(* Logix 5000 project; controller R400_500_XLS vendor 1 type 14 code 216 rev 31.11; software revision 31.01; part 19 of 32 *)
(* tags used below, declared in another part *)
   Alarm : SINT;   // Wait 3 seconds
   Condenser : INT;
   DRYING : DINT;   // Drying id number
   FINAL_RINSE_MAX_NBR : INT;   // Maximum nimber of final rinse
   LowPressAlmSp : REAL;   // Pump pressure too low setpoint
   M : DINT[5];   // Memory Bits
   MaxTrtTempSp : REAL;
   ONS_FC85 : SINT;
   PURE_WATER_HEATING_TIME : DINT;   // Time before an alarm is thrown when the pure water tank is heating
   PWTnkTempAlmSp : REAL;   // Pure water tank temperature too high setpoint
   s00_Nb : STRING;
   s0_Nb : STRING;
   s2lastdigits : STRING;
   s36 : STRING;
   s360 : STRING;
   s3600 : STRING;
   s36000 : STRING;
   s360000 : STRING;
   s3600000 : STRING;
   s36000000 : STRING;
   s360000000 : STRING;
   sDigits1_2 : STRING;
   Service : DINT[2];   // Unused Service Mode Memory Bit
   ServicePassword : DINT;   // Service Password
   sInvertedPairs : STRING;
   sLastdigit : STRING;
   SRE3_Serial_Number : STRING;   // Serial number
   start_1 : SINT;
   start_2 : SINT;
   sTempo1 : STRING;
   sTempo2 : STRING;
   SumpTempAlmSp : REAL;   // Sump temperature too high setpoint
   Tmr : TIMER[107];
   bInibitAutologout : BOOL;   // Cancel AutoLogout
   BoilingValue : REAL;
   Cfg_10_Modules : BOOL;   // Chassis is configured 10 slots
   ChemicalName : STRING[9];   // Used by HMI
   COOLING_PHASE_TIME : DINT;   // Time of the cooling phase when time based drying
   DrainExtensionTime : DINT;
   iDelayBeforeFillingAuthAlarmMM : DINT;
   iDelayBeforeFillingAuthAlarmSS : DINT;
   iInactivityLogoutTime : DINT;   // Inactivity Logout Time In Minutes
   iInactivityPeriod : DINT;   // Inactivity Period before Logout * Value Must be greater than 0
   iPWClosingDelayMM : DINT;
   iPWClosingDelaySS : DINT;
   Non_Vented_with_Dry_Option : BOOL;
   NonVented_Without_Dry_Option : BOOL;
   NumInput : UDT_NUMERIC_INPUT[65];   // Numeric input
   NumInputReal : UDT_NUMERIC_INPUT_REAL[17];
   Screen_Ctrl : DINT;   // PLC Screen Request
   tDelayBeforeFillingAuthAlarm : TIMER;
   tDelayBeforeTankFillingAuthAlarm : TIMER;
   Tpb : DINT[11];
   tPureWaterTankClosingDelay : TIMER;
   tPWClosingDelay : TIMER;
   TRUE : BOOL;   // Always true bit
   Unit : Hrdwre;   // Unit Configuration
   Vented_with_Dry_Option : BOOL;
(* MainProgram, continued *)

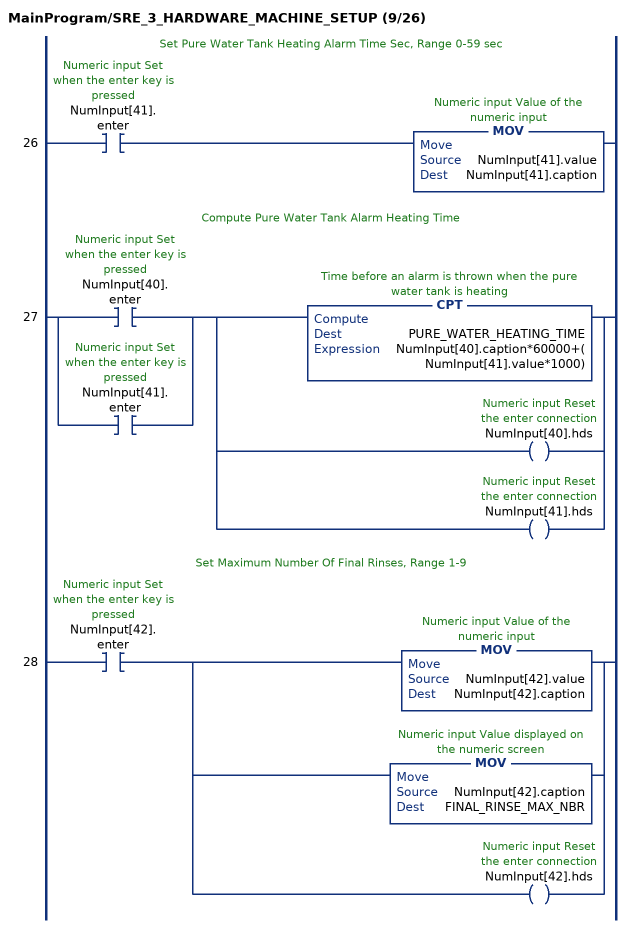
   [picture p363: MainProgram/SRE_3_HARDWARE_MACHINE_SETUP rungs 26-28]
   // Set Pure Water Tank Heating Alarm Time Sec, Range 0-59 sec
   26: XIC(NumInput[41].enter)MOV(NumInput[41].value,NumInput[41].caption);
   // Compute Pure Water Tank Alarm Heating Time
   27: [XIC(NumInput[40].enter) ,XIC(NumInput[41].enter) ][CPT(PURE_WATER_HEATING_TIME,NumInput[40].caption*60000+(NumInput[41].value*1000)) ,OTE(NumInput[40].hds) ,OTE(NumInput[41].hds) ];
   // Set Maximum Number Of Final Rinses, Range 1-9
   28: XIC(NumInput[42].enter)[MOV(NumInput[42].value,NumInput[42].caption) ,MOV(NumInput[42].caption,FINAL_RINSE_MAX_NBR) ,OTE(NumInput[42].hds) ];
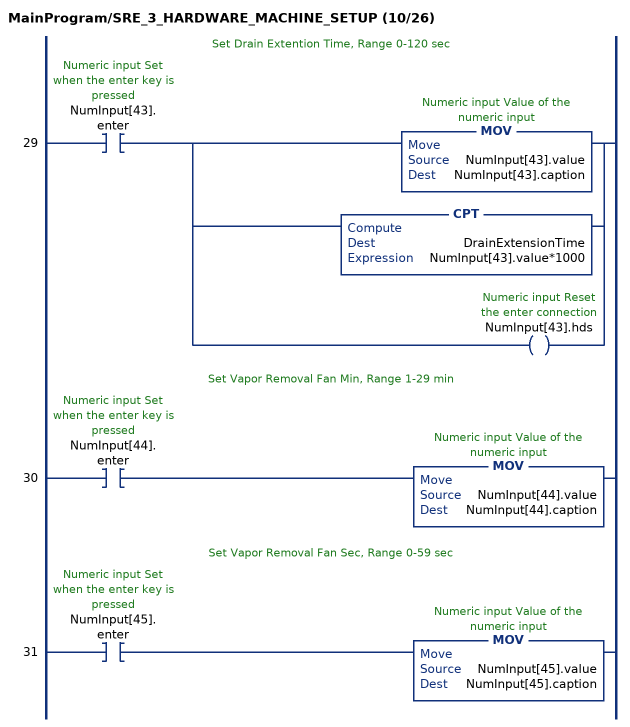
   // Set Drain Extention Time, Range 0-120 sec
   29: XIC(NumInput[43].enter)[MOV(NumInput[43].value,NumInput[43].caption) ,CPT(DrainExtensionTime,NumInput[43].value*1000) ,OTE(NumInput[43].hds) ];
   // Set Vapor Removal Fan Min, Range 1-29 min
   30: XIC(NumInput[44].enter)MOV(NumInput[44].value,NumInput[44].caption);
   // Set Vapor Removal Fan Sec, Range 0-59 sec
   31: XIC(NumInput[45].enter)MOV(NumInput[45].value,NumInput[45].caption);
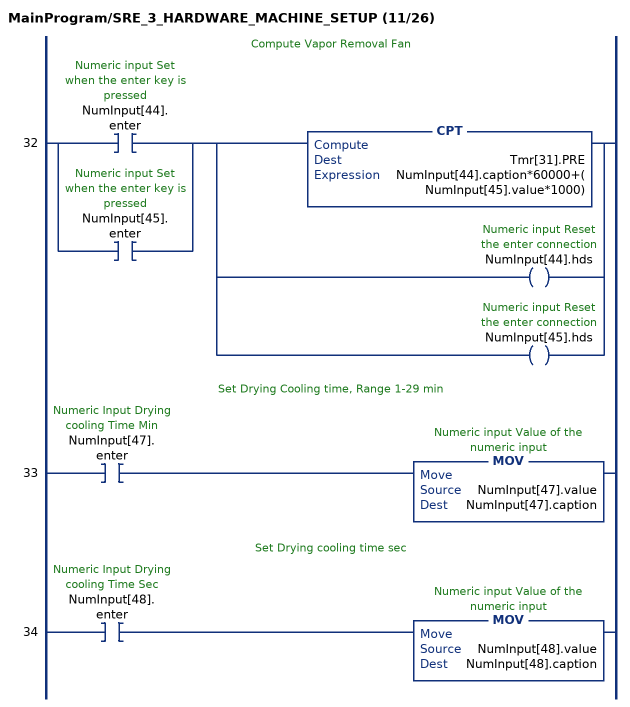
   // Compute Vapor Removal Fan
   32: [XIC(NumInput[44].enter) ,XIC(NumInput[45].enter) ][CPT(Tmr[31].PRE,NumInput[44].caption*60000+(NumInput[45].value*1000)) ,OTE(NumInput[44].hds) ,OTE(NumInput[45].hds) ];
   // Set Drying Cooling time, Range 1-29 min
   33: XIC(NumInput[47].enter)MOV(NumInput[47].value,NumInput[47].caption);
   // Set Drying cooling time sec
   34: XIC(NumInput[48].enter)MOV(NumInput[48].value,NumInput[48].caption);
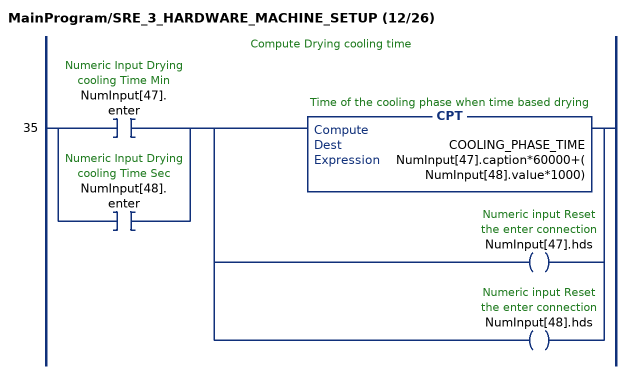
   // Compute Drying cooling time
   35: [XIC(NumInput[47].enter) ,XIC(NumInput[48].enter) ][CPT(COOLING_PHASE_TIME,NumInput[47].caption*60000+(NumInput[48].value*1000)) ,OTE(NumInput[47].hds) ,OTE(NumInput[48].hds) ];
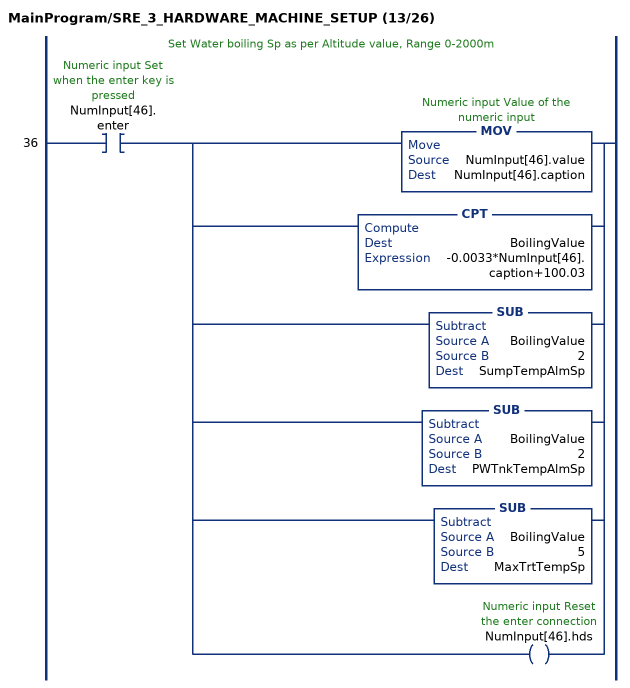
   // Set Water boiling Sp as per Altitude value, Range 0-2000m
   36: XIC(NumInput[46].enter)[MOV(NumInput[46].value,NumInput[46].caption) ,CPT(BoilingValue,-0.0033*NumInput[46].caption+100.03) ,SUB(BoilingValue,2,SumpTempAlmSp) ,SUB(BoilingValue,2,PWTnkTempAlmSp) ,SUB(BoilingValue,5,MaxTrtTempSp) ,OTE(NumInput[46].hds) ];
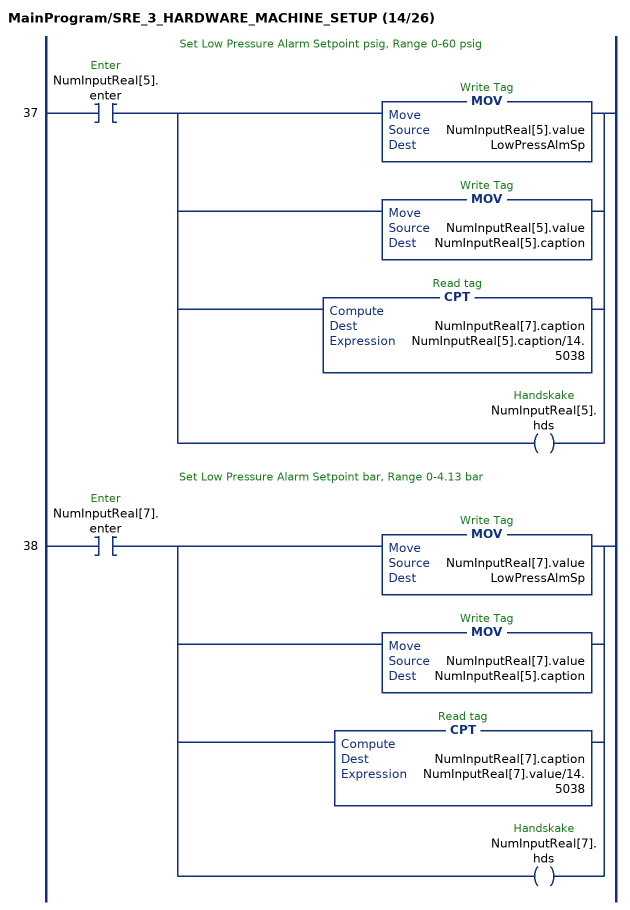
   // Set Low Pressure Alarm Setpoint psig, Range 0-60 psig
   37: XIC(NumInputReal[5].enter)[MOV(NumInputReal[5].value,LowPressAlmSp) ,MOV(NumInputReal[5].value,NumInputReal[5].caption) ,CPT(NumInputReal[7].caption,NumInputReal[5].caption/14.5038) ,OTE(NumInputReal[5].hds) ];
   // Set Low Pressure Alarm Setpoint bar, Range 0-4.13 bar
   38: XIC(NumInputReal[7].enter)[MOV(NumInputReal[7].value,LowPressAlmSp) ,MOV(NumInputReal[7].value,NumInputReal[5].caption) ,CPT(NumInputReal[7].caption,NumInputReal[7].value/14.5038) ,OTE(NumInputReal[7].hds) ];
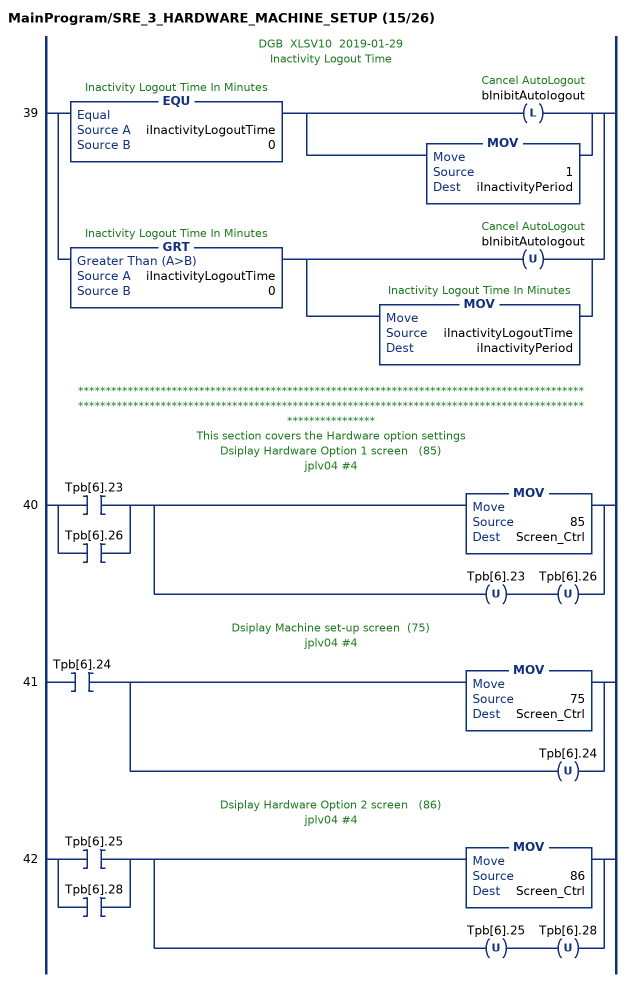
   // DGB  XLSV10  2019-01-29
   // Inactivity Logout Time
   39: [EQU(iInactivityLogoutTime,0) [OTL(bInibitAutologout) ,MOV(1,iInactivityPeriod) ] ,GRT(iInactivityLogoutTime,0) [OTU(bInibitAutologout) ,MOV(iInactivityLogoutTime,iInactivityPeriod) ] ];
   // ********************************************************************************************************************************************************************************************************
   // This section covers the Hardware option settings
   // Dsiplay Hardware Option 1 screen   (85)
   // jplv04 #4
   40: [XIC(Tpb[6].23) ,XIC(Tpb[6].26) ][MOV(85,Screen_Ctrl) ,OTU(Tpb[6].23) OTU(Tpb[6].26) ];
   // Dsiplay Machine set-up screen  (75)
   // jplv04 #4
   41: XIC(Tpb[6].24)[MOV(75,Screen_Ctrl) ,OTU(Tpb[6].24) ];
   // Dsiplay Hardware Option 2 screen   (86)
   // jplv04 #4
   42: [XIC(Tpb[6].25) ,XIC(Tpb[6].28) ][MOV(86,Screen_Ctrl) ,OTU(Tpb[6].25) OTU(Tpb[6].28) ];
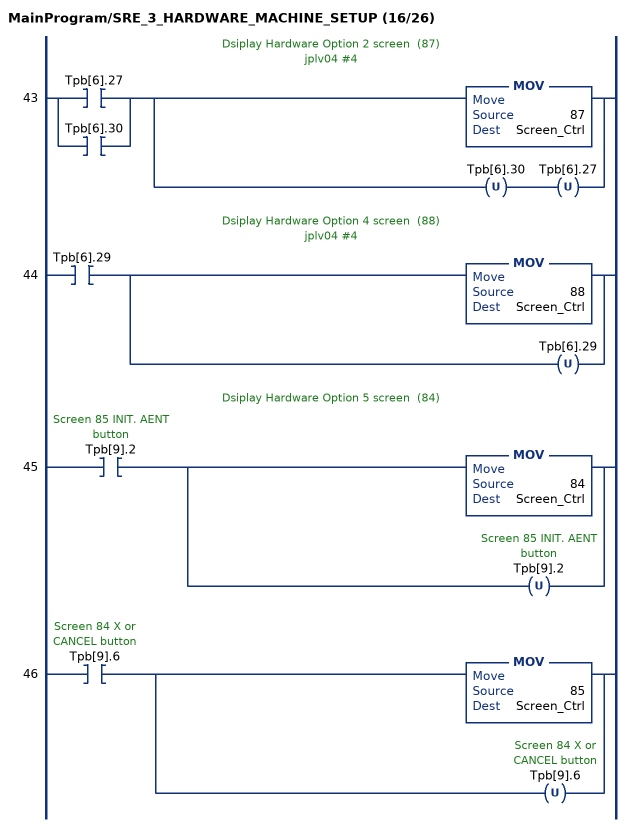
   // Dsiplay Hardware Option 2 screen  (87)
   // jplv04 #4
   43: [XIC(Tpb[6].27) ,XIC(Tpb[6].30) ][MOV(87,Screen_Ctrl) ,OTU(Tpb[6].30) OTU(Tpb[6].27) ];
   // Dsiplay Hardware Option 4 screen  (88)
   // jplv04 #4
   44: XIC(Tpb[6].29)[MOV(88,Screen_Ctrl) ,OTU(Tpb[6].29) ];
   // Dsiplay Hardware Option 5 screen  (84)
   45: XIC(Tpb[9].2)[MOV(84,Screen_Ctrl) ,OTU(Tpb[9].2) ];
   46: XIC(Tpb[9].6)[MOV(85,Screen_Ctrl) ,OTU(Tpb[9].6) ];
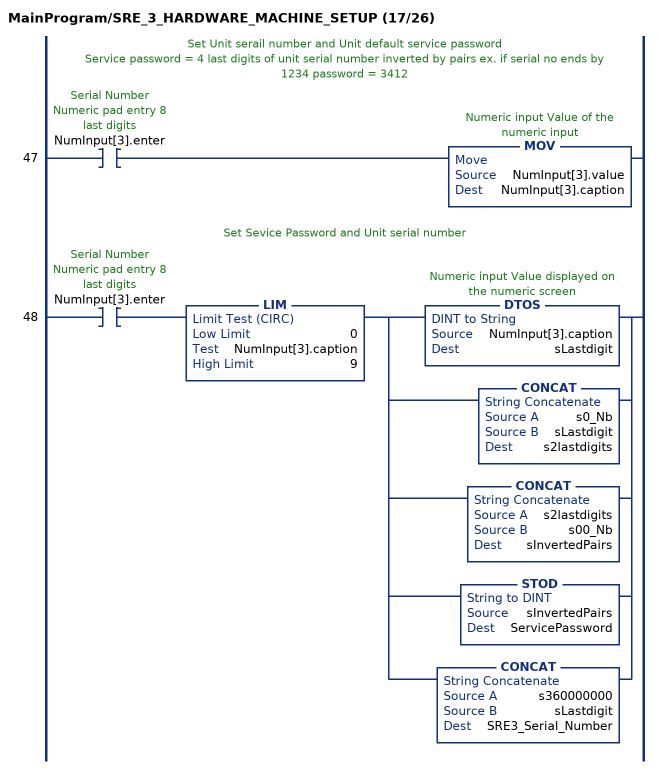
   // Set Unit serail number and Unit default service password
   // Service password = 4 last digits of unit serial number inverted by pairs ex. if serial no ends by 1234 password = 3412
   47: XIC(NumInput[3].enter)MOV(NumInput[3].value,NumInput[3].caption);
   // Set Sevice Password and Unit serial number
   48: XIC(NumInput[3].enter)LIM(0,NumInput[3].caption,9)[DTOS(NumInput[3].caption,sLastdigit) ,CONCAT(s0_Nb,sLastdigit,s2lastdigits) ,CONCAT(s2lastdigits,s00_Nb,sInvertedPairs) ,STOD(sInvertedPairs,ServicePassword) ,CONCAT(s360000000,sLastdigit,SRE3_Serial_Number) ];
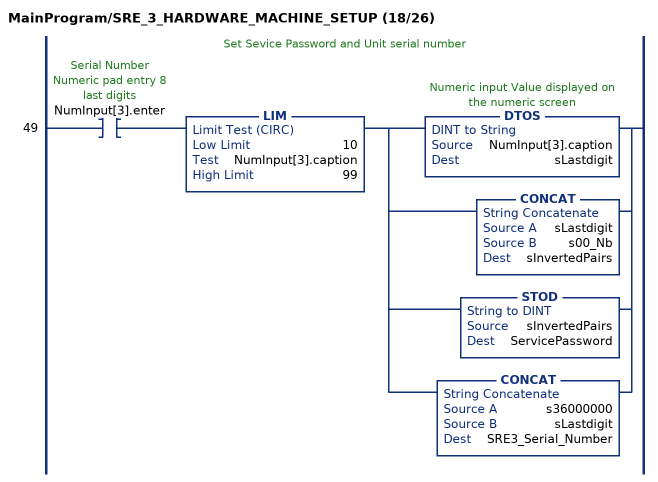
   // Set Sevice Password and Unit serial number
   49: XIC(NumInput[3].enter)LIM(10,NumInput[3].caption,99)[DTOS(NumInput[3].caption,sLastdigit) ,CONCAT(sLastdigit,s00_Nb,sInvertedPairs) ,STOD(sInvertedPairs,ServicePassword) ,CONCAT(s36000000,sLastdigit,SRE3_Serial_Number) ];
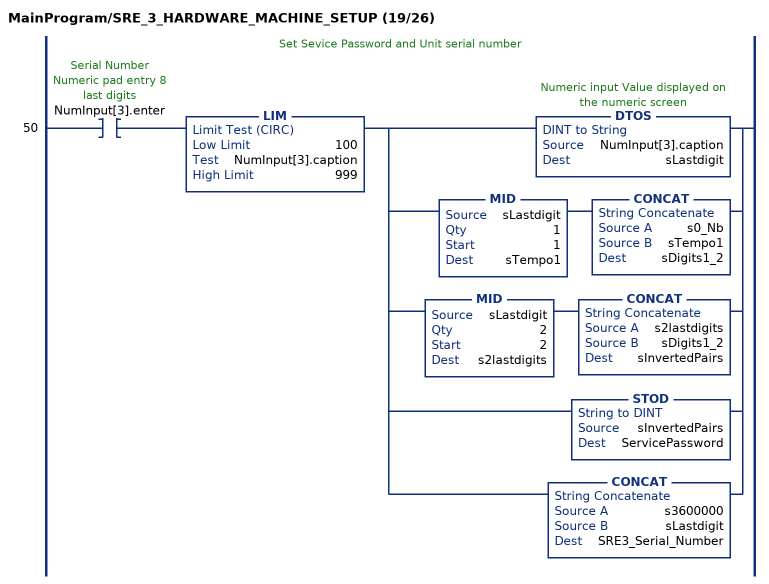
   // Set Sevice Password and Unit serial number
   50: XIC(NumInput[3].enter)LIM(100,NumInput[3].caption,999)[DTOS(NumInput[3].caption,sLastdigit) ,MID(sLastdigit,1,1,sTempo1) CONCAT(s0_Nb,sTempo1,sDigits1_2) ,MID(sLastdigit,2,2,s2lastdigits) CONCAT(s2lastdigits,sDigits1_2,sInvertedPairs) ,STOD(sInvertedPairs,ServicePassword) ,CONCAT(s3600000,sLastdigit,SRE3_Serial_Number) ];
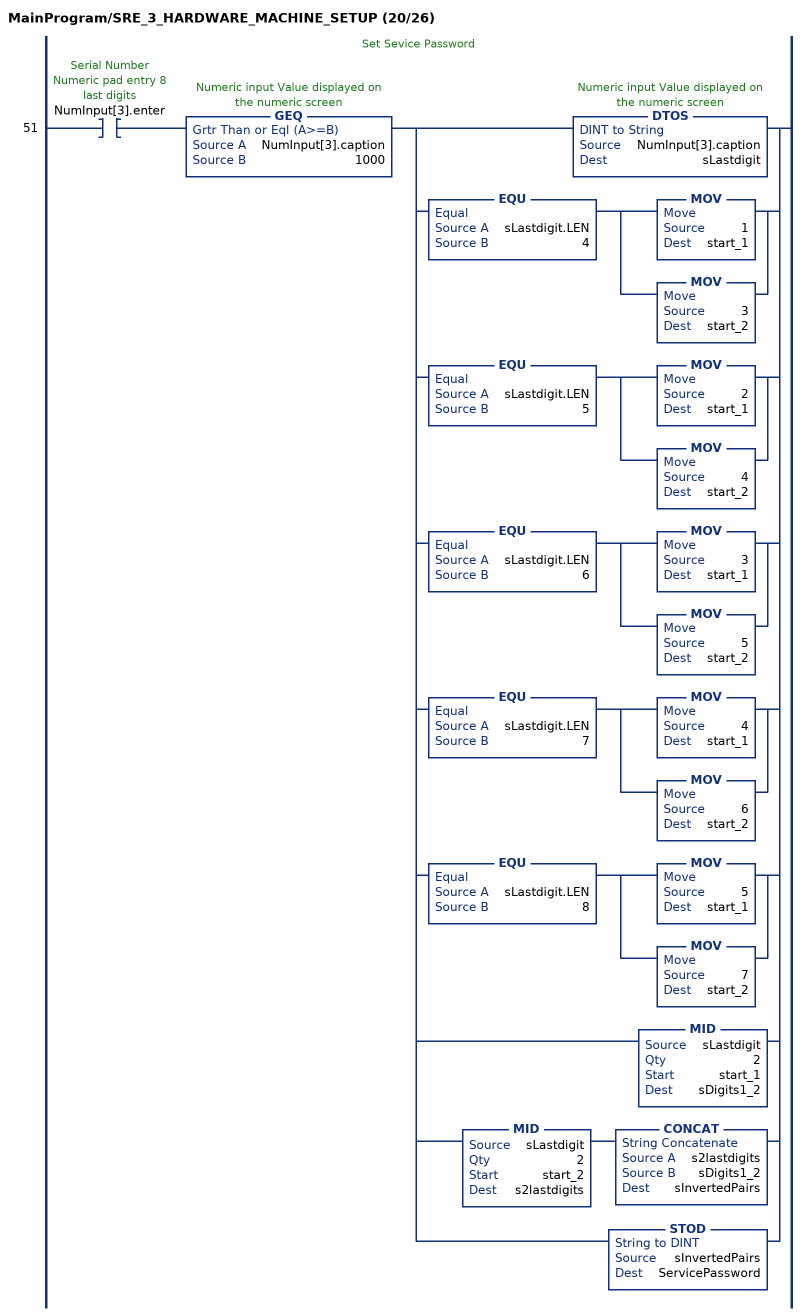
   // Set Sevice Password
   51: XIC(NumInput[3].enter)GEQ(NumInput[3].caption,1000)[DTOS(NumInput[3].caption,sLastdigit) ,EQU(sLastdigit.LEN,4) [MOV(1,start_1) ,MOV(3,start_2) ] ,EQU(sLastdigit.LEN,5) [MOV(2,start_1) ,MOV(4,start_2) ] ,EQU(sLastdigit.LEN,6) [MOV(3,start_1) ,MOV(5,start_2) ] ,EQU(sLastdigit.LEN,7) [MOV(4,start_1) ,MOV(6,start_2) ] ,EQU(sLastdigit.LEN,8) [MOV(5,start_1) ,MOV(7,start_2) ] ,MID(sLastdigit,2,start_1,sDigits1_2) ,MID(sLastdigit,2,start_2,s2lastdigits) CONCAT(s2lastdigits,sDigits1_2,sInvertedPairs) ,STOD(sInvertedPairs,ServicePassword) ];
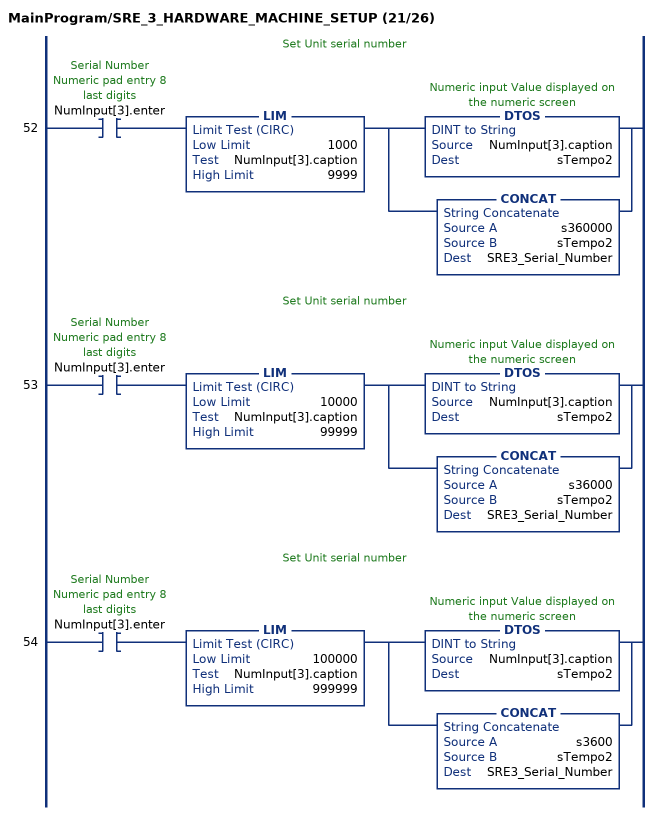
   // Set Unit serial number
   52: XIC(NumInput[3].enter)LIM(1000,NumInput[3].caption,9999)[DTOS(NumInput[3].caption,sTempo2) ,CONCAT(s360000,sTempo2,SRE3_Serial_Number) ];
   // Set Unit serial number
   53: XIC(NumInput[3].enter)LIM(10000,NumInput[3].caption,99999)[DTOS(NumInput[3].caption,sTempo2) ,CONCAT(s36000,sTempo2,SRE3_Serial_Number) ];
   // Set Unit serial number
   54: XIC(NumInput[3].enter)LIM(100000,NumInput[3].caption,999999)[DTOS(NumInput[3].caption,sTempo2) ,CONCAT(s3600,sTempo2,SRE3_Serial_Number) ];
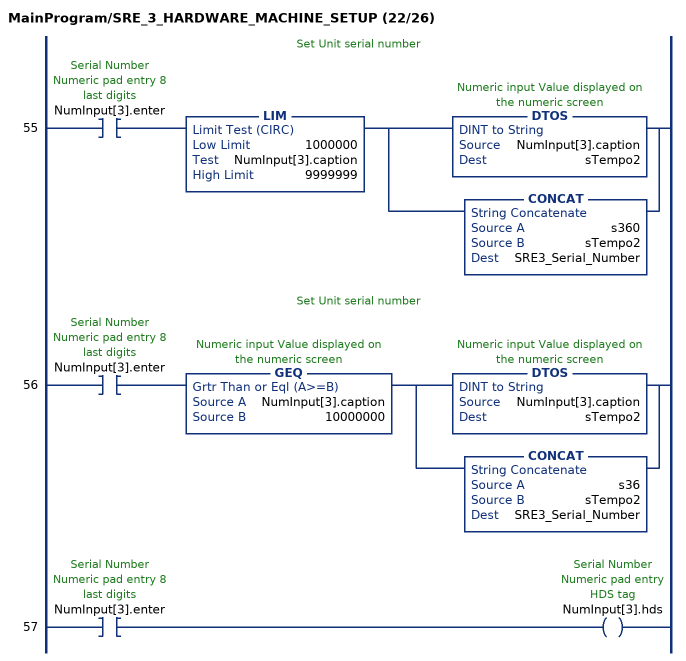
   // Set Unit serial number
   55: XIC(NumInput[3].enter)LIM(1000000,NumInput[3].caption,9999999)[DTOS(NumInput[3].caption,sTempo2) ,CONCAT(s360,sTempo2,SRE3_Serial_Number) ];
   // Set Unit serial number
   56: XIC(NumInput[3].enter)GEQ(NumInput[3].caption,10000000)[DTOS(NumInput[3].caption,sTempo2) ,CONCAT(s36,sTempo2,SRE3_Serial_Number) ];
   57: XIC(NumInput[3].enter)OTE(NumInput[3].hds);
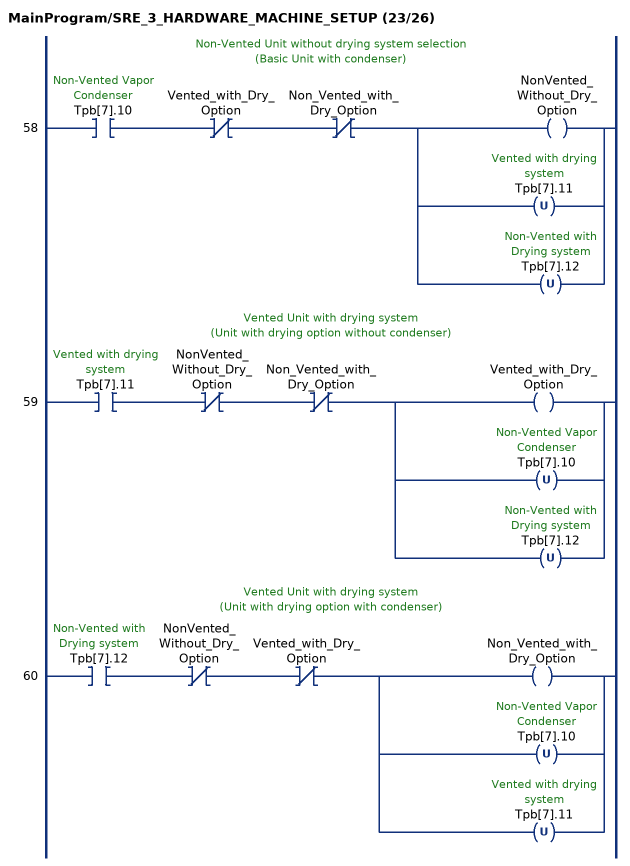
   // Non-Vented Unit without drying system selection
   // (Basic Unit with condenser)
   58: XIC(Tpb[7].10)XIO(Vented_with_Dry_Option)XIO(Non_Vented_with_Dry_Option)[OTE(NonVented_Without_Dry_Option) ,OTU(Tpb[7].11) ,OTU(Tpb[7].12) ];
   // Vented Unit with drying system
   // (Unit with drying option without condenser)
   59: XIC(Tpb[7].11)XIO(NonVented_Without_Dry_Option)XIO(Non_Vented_with_Dry_Option)[OTE(Vented_with_Dry_Option) ,OTU(Tpb[7].10) ,OTU(Tpb[7].12) ];
   // Vented Unit with drying system
   // (Unit with drying option with condenser)
   60: XIC(Tpb[7].12)XIO(NonVented_Without_Dry_Option)XIO(Vented_with_Dry_Option)[OTE(Non_Vented_with_Dry_Option) ,OTU(Tpb[7].10) ,OTU(Tpb[7].11) ];
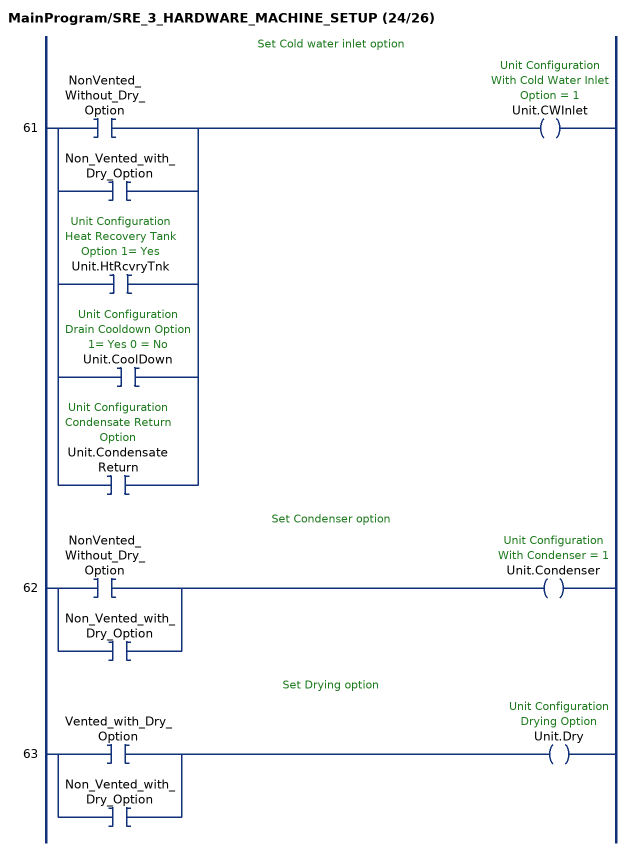
   // Set Cold water inlet option
   61: [XIC(NonVented_Without_Dry_Option) ,XIC(Non_Vented_with_Dry_Option) ,XIC(Unit.HtRcvryTnk) ,XIC(Unit.CoolDown) ,XIC(Unit.CondensateReturn) ]OTE(Unit.CWInlet);
   // Set Condenser option
   62: [XIC(NonVented_Without_Dry_Option) ,XIC(Non_Vented_with_Dry_Option) ]OTE(Unit.Condenser);
   // Set Drying option
   63: [XIC(Vented_with_Dry_Option) ,XIC(Non_Vented_with_Dry_Option) ]OTE(Unit.Dry);
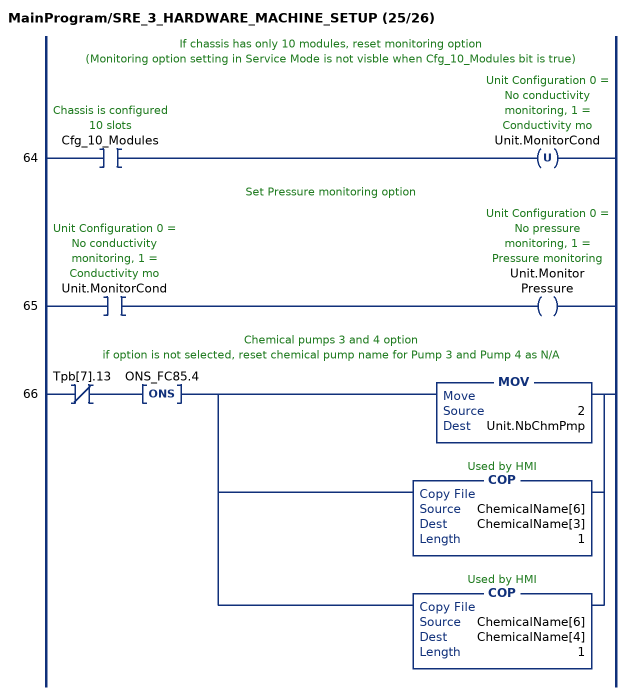
   // If chassis has only 10 modules, reset monitoring option
   // (Monitoring option setting in Service Mode is not visble when Cfg_10_Modules bit is true)
   64: XIC(Cfg_10_Modules)OTU(Unit.MonitorCond);
   // Set Pressure monitoring option
   65: XIC(Unit.MonitorCond)OTE(Unit.MonitorPressure);
   // Chemical pumps 3 and 4 option
   // if option is not selected, reset chemical pump name for Pump 3 and Pump 4 as N/A
   66: XIO(Tpb[7].13)ONS(ONS_FC85.4)[MOV(2,Unit.NbChmPmp) ,COP(ChemicalName[6],ChemicalName[3],1) ,COP(ChemicalName[6],ChemicalName[4],1) ];
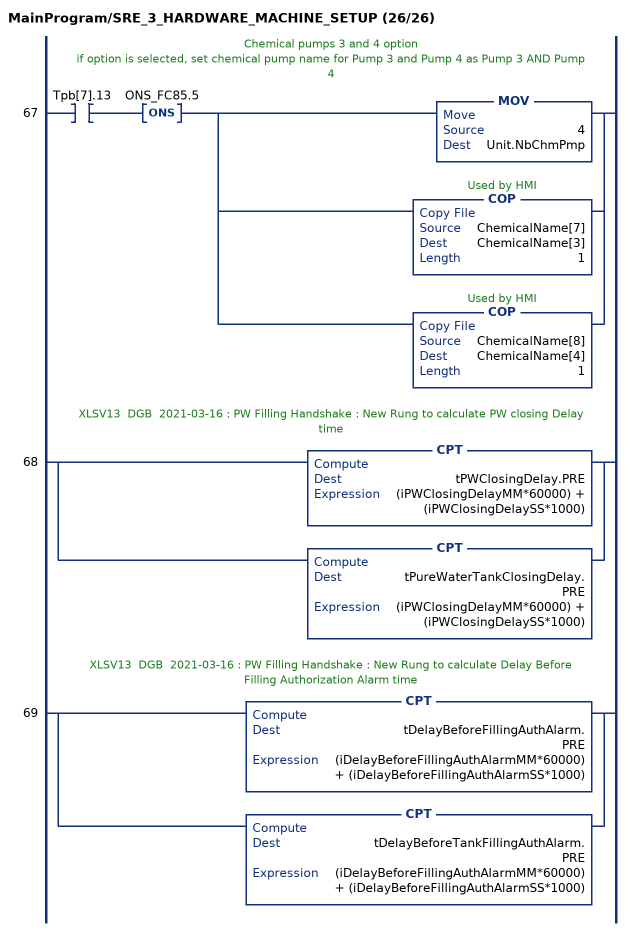
   // Chemical pumps 3 and 4 option
   // if option is selected, set chemical pump name for Pump 3 and Pump 4 as Pump 3 AND Pump 4
   67: XIC(Tpb[7].13)ONS(ONS_FC85.5)[MOV(4,Unit.NbChmPmp) ,COP(ChemicalName[7],ChemicalName[3],1) ,COP(ChemicalName[8],ChemicalName[4],1) ];
   // XLSV13  DGB  2021-03-16 : PW Filling Handshake : New Rung to calculate PW closing Delay time
   68: [CPT(tPWClosingDelay.PRE,(iPWClosingDelayMM*60000) + (iPWClosingDelaySS*1000)) ,CPT(tPureWaterTankClosingDelay.PRE,(iPWClosingDelayMM*60000) + (iPWClosingDelaySS*1000)) ];
   // XLSV13  DGB  2021-03-16 : PW Filling Handshake : New Rung to calculate Delay Before Filling Authorization Alarm time
   69: [CPT(tDelayBeforeFillingAuthAlarm.PRE,(iDelayBeforeFillingAuthAlarmMM*60000) + (iDelayBeforeFillingAuthAlarmSS*1000)) ,CPT(tDelayBeforeTankFillingAuthAlarm.PRE,(iDelayBeforeFillingAuthAlarmMM*60000) + (iDelayBeforeFillingAuthAlarmSS*1000)) ];
END_ROUTINE
